(* IEC 61131-3 sources: ZPLC/tools/hil/st_tests, 25 files *)

(* ---- full_language_test.st ---- *)
TYPE State : (INIT, PROCESS, DONE, ERROR); END_TYPE

FUNCTION_BLOCK FB_Logger
    VAR
        LastMsg : WSTRING;
        MsgCount : INT := 0;
    END_VAR

    METHOD PUBLIC Log : BOOL
        VAR_INPUT
            Msg : WSTRING;
        END_VAR
        THIS.LastMsg := Msg;
        THIS.MsgCount := THIS.MsgCount + 1;
        Log := TRUE;
    END_METHOD
END_FUNCTION_BLOCK

FUNCTION_BLOCK FB_Process EXTENDS FB_Logger
    VAR
        Timestamp : DT;
        Result : REAL;
    END_VAR

    METHOD PUBLIC Calc : REAL
        VAR_INPUT
            InVal : REAL;
        END_VAR
        VAR_TEMP
            tmp : REAL;
        END_VAR

        tmp := tmp + InVal * 2.0;
        Calc := tmp;
    END_METHOD
END_FUNCTION_BLOCK

PROGRAM FullTest
    VAR
        machine : FB_Process;
        currentState : State := INIT;

        test_dt : DT;
        calc_res1 AT %QD1 : REAL;
        calc_res2 AT %QD2 : REAL;

        cycle AT %QW0 : INT := 0;

        flag_enum AT %QX12.0 : BOOL;
        flag_oop AT %QX12.1 : BOOL;
        flag_temp AT %QX12.2 : BOOL;
        flag_types AT %QX12.3 : BOOL;
    END_VAR

    cycle := cycle + 1;

    CASE currentState OF
        0: (* INIT *)
            machine.Log(Msg := "Start");
            machine.Timestamp := DT#2024-01-01-12:00:00;
            test_dt := machine.Timestamp;
            currentState := 1;

        1: (* PROCESS *)
            calc_res1 := machine.Calc(InVal := 10.0);
            calc_res2 := machine.Calc(InVal := 20.0);
            currentState := 2;

        2: (* DONE *)
            flag_enum := TRUE;

            IF machine.MsgCount = 1 THEN flag_oop := TRUE; END_IF;

            IF calc_res1 = 20.0 AND calc_res2 = 40.0 THEN flag_temp := TRUE; END_IF;

            IF test_dt > DT#2023-01-01-00:00:00 THEN flag_types := TRUE; END_IF;
    END_CASE;

END_PROGRAM

(* ---- named_params_test.st ---- *)
FUNCTION_BLOCK FB_Calc
    METHOD PUBLIC Add : REAL
        VAR_INPUT
            A : REAL;
            B : REAL;
        END_VAR
        Add := A + B;
    END_METHOD
END_FUNCTION_BLOCK

PROGRAM NamedParamsTest
    VAR
        calc : FB_Calc;
        res AT %QD0 : REAL;
    END_VAR

    res := calc.Add(A := 10.0, B := 20.0);
END_PROGRAM

(* ---- oop_extends.st ---- *)
FUNCTION_BLOCK FB_Base
VAR
    BaseVal : INT;
END_VAR

METHOD PUBLIC InitBase : BOOL
    THIS.BaseVal := 10;
    InitBase := TRUE;
END_METHOD

METHOD PUBLIC GetBase : INT
    GetBase := THIS.BaseVal;
END_METHOD

METHOD PUBLIC VirtualMethod : INT
    VirtualMethod := 111;
END_METHOD
END_FUNCTION_BLOCK

FUNCTION_BLOCK FB_Child EXTENDS FB_Base
VAR
    ChildVal : INT;
END_VAR

METHOD PUBLIC InitChild : BOOL
    THIS.BaseVal := 10;
    THIS.ChildVal := 20;
    InitChild := TRUE;
END_METHOD

METHOD PUBLIC GetChild : INT
    GetChild := THIS.ChildVal;
END_METHOD

METHOD PUBLIC OVERRIDE VirtualMethod : INT
    VirtualMethod := 222;
END_METHOD
END_FUNCTION_BLOCK

PROGRAM TestExtends
VAR
    base : FB_Base;
    child : FB_Child;

    res_base_base : INT;
    res_child_base : INT;
    res_child_child : INT;
    res_virt_base : INT;
    res_virt_child : INT;

    initialized : BOOL := FALSE;
    dummy : BOOL;

    test_passed AT %QX0.0 : BOOL := FALSE;
    debug_val AT %QW1 : INT;
    life_counter AT %QW2 : INT; (* 0x1004 *)
END_VAR

life_counter := life_counter + 1;

IF NOT initialized THEN
    dummy := base.InitBase();
    dummy := child.InitChild();
    initialized := TRUE;
END_IF;

res_base_base := base.GetBase();
res_child_base := child.GetBase();
res_child_child := child.GetChild();

res_virt_base := base.VirtualMethod();
res_virt_child := child.VirtualMethod();

debug_val := res_virt_child;

IF res_base_base = 10 AND
   res_child_base = 10 AND
   res_child_child = 20 AND
   res_virt_base = 111 AND
   res_virt_child = 222 THEN
    test_passed := TRUE;
END_IF;

END_PROGRAM

(* ---- oop_extends_simple.st ---- *)
FUNCTION_BLOCK FB_Base
METHOD PUBLIC GetVal : INT
    GetVal := 111;
END_METHOD
END_FUNCTION_BLOCK

FUNCTION_BLOCK FB_Child EXTENDS FB_Base
METHOD PUBLIC OVERRIDE GetVal : INT
    GetVal := 222;
END_METHOD
END_FUNCTION_BLOCK

PROGRAM SimpleExtends
VAR
    child : FB_Child;
    res : INT;
    debug AT %QW0 : INT;
END_VAR

res := child.GetVal();
debug := res;
END_PROGRAM

(* ---- oop_test.st ---- *)
(*
 * ZPLC OOP HIL Test
 *
 * Tests IEC 61131-3 OOP extensions:
 * - FUNCTION_BLOCK with METHOD
 * - THIS keyword
 * - Method calls on FB instances
 *
 * Memory Layout (OPI starts at 0x1000):
 * - 0x1000: test_passed BOOL
 * - 0x1002: counter_value INT (2 bytes)
 * - 0x1004: method_result INT (2 bytes)
 * - 0x1006: cycle_count INT (2 bytes)
 *)

(* Simple Counter FB with Methods *)
FUNCTION_BLOCK FB_Counter
VAR
    Count : INT;
    MaxVal : INT;
END_VAR

(* Reset counter to zero *)
METHOD PUBLIC Reset : BOOL
    THIS.Count := 0;
    THIS.MaxVal := 100;
    Reset := TRUE;
END_METHOD

(* Increment counter by 1 and return new value *)
METHOD PUBLIC Increment : INT
    THIS.Count := THIS.Count + 1;
    Increment := THIS.Count;
END_METHOD

(* Get current count value *)
METHOD PUBLIC GetValue : INT
    GetValue := THIS.Count;
END_METHOD

(* Add 10 to counter *)
METHOD PUBLIC AddTen : INT
    THIS.Count := THIS.Count + 10;
    AddTen := THIS.Count;
END_METHOD

END_FUNCTION_BLOCK

PROGRAM OOPTest
VAR
    (* Output mappings for test verification *)
    test_passed AT %QX0.0 : BOOL := FALSE;  (* 0x1000 bit 0 *)
    counter_value AT %QW1 : INT;            (* 0x1002 *)
    method_result AT %QW2 : INT;            (* 0x1004 *)
    cycle_count AT %QW3 : INT;              (* 0x1006 *)

    (* FB instance *)
    myCounter : FB_Counter;

    (* Local variables *)
    initialized : BOOL := FALSE;
    temp : INT;
    cycles : INT := 0;
END_VAR

(* Increment cycle counter *)
cycles := cycles + 1;
cycle_count := cycles;

(* Only run initialization once *)
IF NOT initialized THEN
    (* Reset counter to zero *)
    myCounter.Reset();
    initialized := TRUE;
END_IF;

(* Each cycle: increment, then add 10 *)
(* Cycle 1: 0 -> 1 -> 11 *)
(* Cycle 2: 11 -> 12 -> 22 *)

temp := myCounter.Increment();
method_result := myCounter.AddTen();
counter_value := myCounter.GetValue();

(* Test passes if counter >= 11 (at least one full cycle completed) *)
IF counter_value >= 11 THEN
    test_passed := TRUE;
END_IF;

END_PROGRAM

(* ---- user_fb.st ---- *)
FUNCTION_BLOCK MyCounter
VAR_INPUT
    Up : BOOL;
END_VAR
VAR_OUTPUT
    Count : INT := 0;
END_VAR
VAR
    prev_up : BOOL := FALSE;
END_VAR

    (* Rising Edge Detection *)
    IF Up AND NOT prev_up THEN
        Count := Count + 1;
    END_IF;
    prev_up := Up;

END_FUNCTION_BLOCK

PROGRAM UserFBTest
VAR
    c1 : MyCounter;
    clk : BOOL := FALSE;
    res_count AT %QW0 : INT; (* 0x1000 *)

    cycle : INT := 0;
END_VAR

cycle := cycle + 1;

(* Generate pulse every 2 cycles: 0->F, 1->F, 2->T, 3->F, 4->T ... *)
clk := (cycle MOD 2) = 0;

c1(Up := clk);
res_count := c1.Count;

END_PROGRAM

(* ---- vartemp_hil.st ---- *)
FUNCTION_BLOCK FB_TempTest
    METHOD PUBLIC AddTemp : INT
        VAR_INPUT In : INT; END_VAR
        VAR_TEMP tmp : INT := 0; END_VAR

        (* tmp should be 0 at start of every call *)
        tmp := tmp + In;
        AddTemp := tmp;
    END_METHOD
END_FUNCTION_BLOCK

PROGRAM Main
    VAR
        fb : FB_TempTest;
        res1 AT %QW0 : INT;
        res2 AT %QW1 : INT;
    END_VAR

    res1 := fb.AddTemp(In := 10);
    res2 := fb.AddTemp(In := 20);
END_PROGRAM

(* ---- complex_types.st ---- *)
PROGRAM ComplexTypes
VAR
    matrix : ARRAY[0..1, 0..1] OF INT;
    sum : INT;

    (* Result on the output image, byte 0 (0x1000) *)
    res_x AT %QW0 : INT;
END_VAR

(* Initialize Matrix *)
matrix[0,0] := 10;
matrix[0,1] := 20;
matrix[1,0] := 30;
matrix[1,1] := 40;

(* Calculate diagonal sum: 10 + 40 = 50 *)
sum := matrix[0,0] + matrix[1,1];

(* Output *)
res_x := sum;

END_PROGRAM

(* ---- counters_extra.st ---- *)
PROGRAM TestCounters
VAR
    (* CTD Test *)
    myCtd : CTD;
    cd : BOOL;
    ld : BOOL;
    pv : INT := 5;
    q_ctd AT %QX0.0 : BOOL;
    cv_ctd AT %QW1 : INT;

    (* CTUD Test *)
    myCtud : CTUD;
    cu : BOOL;
    cd_ud : BOOL;
    r : BOOL;
    ld_ud : BOOL;
    pv_ud : INT := 5;
    qu AT %QX0.1 : BOOL;
    qd AT %QX0.2 : BOOL;
    cv_ud AT %QW2 : INT;

    step : INT := 0;
    cycles : INT := 0;
END_VAR

cycles := cycles + 1;

(* State Machine to generate edges *)
CASE step OF
    0: (* Init *)
        ld := TRUE; (* CTD: Load 5 *)
        r := TRUE;  (* CTUD: Reset to 0 *)
        step := 1;

    1: (* Release controls *)
        ld := FALSE;
        r := FALSE;
        step := 2;

    2: (* Generate 3 down pulses for CTD *)
        cd := TRUE;
        step := 3;
    3:
        cd := FALSE;
        step := 4;
    4:
        cd := TRUE;
        step := 5;
    5:
        cd := FALSE;
        step := 6;
    6:
        cd := TRUE;
        step := 7;
    7:
        cd := FALSE;
        (* CTD started at 5. 3 pulses -> 2. *)

        (* Generate 6 up pulses for CTUD *)
        cu := TRUE;
        step := 8;
    8:
        cu := FALSE;
        (* Repeat up to 6 times using modulo logic or just linear steps *)
        IF cycles > 30 THEN
            step := 99;
        ELSE
            (* Toggle CU every even/odd step *)
            IF (cycles MOD 2) = 0 THEN cu := TRUE; ELSE cu := FALSE; END_IF;
        END_IF;

    99: (* Done *)
        cu := FALSE;
        cd := FALSE;
END_CASE;

(* Call FBs *)
myCtd(CD := cd, LD := ld, PV := pv);
q_ctd := myCtd.Q;
cv_ctd := myCtd.CV;

myCtud(CU := cu, CD := cd_ud, R := r, LD := ld_ud, PV := pv_ud);
qu := myCtud.QU;
qd := myCtud.QD;
cv_ud := myCtud.CV;

END_PROGRAM

(* ---- loop_control.st ---- *)
PROGRAM LoopControl
VAR
    i : INT;
    j : INT;
    sum : INT := 0;

    res_exit AT %QW0 : INT;    (* 0x1000 *)
    res_cont AT %QW1 : INT;    (* 0x1002 *)
END_VAR

(* EXIT Test: Stop at 5 *)
FOR i := 1 TO 10 DO
    IF i = 5 THEN
        EXIT;
    END_IF;
END_FOR;
res_exit := i;

(* CONTINUE Test: Sum all except 3 (1+2+4+5=12) *)
sum := 0;
FOR j := 1 TO 5 DO
    IF j = 3 THEN
        CONTINUE;
    END_IF;
    sum := sum + j;
END_FOR;
res_cont := sum;

END_PROGRAM

(* ---- loop_test.st ---- *)
PROGRAM LoopTest
VAR
    i : INT := 0;
    j : INT := 0;

    res_while AT %QW0 : INT;  (* 0x1000 *)
    res_repeat AT %QW1 : INT; (* 0x1002 *)
END_VAR

(* WHILE Loop *)
WHILE i < 10 DO
    i := i + 1;
END_WHILE;
res_while := i;

(* REPEAT Loop *)
REPEAT
    j := j + 1;
UNTIL j = 20
END_REPEAT;
res_repeat := j;

(* Reset for next cycle *)
IF i >= 10 THEN i := 0; END_IF;
IF j >= 20 THEN j := 0; END_IF;

END_PROGRAM

(* ---- master_blinky.st ---- *)
PROGRAM MasterBlinky
VAR
    fast_tmr : TON;
    slow_tmr : TON;

    fast_state AT %QX0.1 : BOOL; (* GP1 *)
    slow_state AT %QX0.0 : BOOL; (* GP0 *)

    cycle_count : INT := 0;
END_VAR

(* Fast Blinky (100ms ON / 100ms OFF) *)
fast_tmr(IN := NOT fast_tmr.Q, PT := T#100ms);
IF fast_tmr.Q THEN
    fast_state := NOT fast_state;
END_IF;

(* Slow Blinky (500ms ON / 500ms OFF) *)
slow_tmr(IN := NOT slow_tmr.Q, PT := T#500ms);
IF slow_tmr.Q THEN
    slow_state := NOT slow_state;
END_IF;

cycle_count := cycle_count + 1;

END_PROGRAM

(* ---- master_math_control.st ---- *)
PROGRAM MathControlTest
VAR
    (* Math Results *)
    res_sqrt AT %QD1 : REAL;   (* 0x1004 *)
    res_ln AT %QD2 : REAL;     (* 0x1008 *)
    res_sin AT %QD3 : REAL;   (* 0x100C *)
    res_expt AT %QW8 : INT;   (* 0x1010 *)

    (* Control Results *)
    res_for AT %QW9 : INT;    (* 0x1012 *)
    res_case AT %QW10 : INT;   (* 0x1014 *)

    (* Internal vars *)
    i : INT;
    temp_sum : INT := 0;
    case_sel : INT := 2;
END_VAR

(* 1. Math Tests *)
res_sqrt := SQRT(2.0);
res_ln := LN(2.7182818);
res_sin := SIN(1.570796);
res_expt := REAL_TO_INT(EXPT(2.0, 8));

(* 2. FOR loop test *)
temp_sum := 0;
FOR i := 1 TO 10 DO
    temp_sum := temp_sum + i;
END_FOR;
res_for := temp_sum;

(* 3. CASE test *)
CASE case_sel OF
    1: res_case := 10;
    2: res_case := 20;
    3: res_case := 30;
ELSE
    res_case := 99;
END_CASE;

END_PROGRAM

(* ---- master_test.st ---- *)
PROGRAM MasterTest
VAR
    test_cycle : INT := 0;
    latch_rs : RS;
    latch_sr : SR;
    trig_r : R_TRIG;
    counter : CTU;

    res_rs AT %QX0.0 : BOOL;
    res_sr AT %QX0.1 : BOOL;
    res_trig AT %QX0.2 : BOOL;
    res_ctu AT %QX0.3 : BOOL;
END_VAR

test_cycle := test_cycle + 1;

(* 1. Test RS: Set once and keep it *)
latch_rs(S := (test_cycle = 5), R1 := FALSE);
res_rs := latch_rs.Q1;

(* 2. Test SR: Set once and keep it *)
latch_sr(S1 := (test_cycle = 5), R := FALSE);
res_sr := latch_sr.Q1;

(* 3. Test Trigger: Pulse and latch the result *)
trig_r(CLK := (test_cycle = 5));
IF trig_r.Q THEN
    res_trig := TRUE;
END_IF;

(* 4. Test Counter: Count to 5 and stay there *)
counter(CU := (test_cycle <= 10 AND (test_cycle MOD 2 = 0)), PV := 5, R := (test_cycle = 1));
res_ctu := counter.Q;

END_PROGRAM

(* ---- master_test_2.st ---- *)
PROGRAM MasterTest2
VAR
    test_cycle : INT := 0;
    timer_off : TOF;
    timer_pulse : TP;
    i : INT;
    sum : INT := 0;
    case_val : INT := 0;

    (* Results on the output image: STOP puts the outputs in their safe state, so they are read while it runs *)
    res_tof AT %QX0.0 : BOOL;
    res_tp AT %QX0.1 : BOOL;
    res_for AT %QW1 : INT;
    res_case AT %QW2 : INT;
END_VAR

test_cycle := test_cycle + 1;

timer_off(IN := (test_cycle = 5), PT := T#500ms);
IF test_cycle = 10 AND timer_off.Q THEN
    res_tof := TRUE;
END_IF;

timer_pulse(IN := (test_cycle = 5), PT := T#500ms);
IF test_cycle = 7 AND timer_pulse.Q THEN
    res_tp := TRUE;
END_IF;

IF test_cycle = 10 THEN
    sum := 0;
    FOR i := 1 TO 5 DO
        sum := sum + i;
    END_FOR;
    res_for := sum;
END_IF;

IF test_cycle = 10 THEN
    case_val := 2;
    CASE case_val OF
        1: res_case := 100;
        2: res_case := 200;
    ELSE
        res_case := 0;
    END_CASE;
END_IF;

END_PROGRAM

(* ---- math_real.st ---- *)
PROGRAM MathReal
VAR
    angles : ARRAY[0..2] OF REAL;
    sines : ARRAY[0..2] OF REAL;
    i : INT;

    (* OPI Layout: *)
    (* 0x1000: result_ok (INT, 2 bytes) *)
    (* 0x1004: debug_val (REAL, 4 bytes) *)

    result_ok AT %QW0 : INT;
    debug_val AT %QD1 : REAL;
END_VAR

angles[0] := 0.0;
angles[1] := 1.570796;
angles[2] := 3.141592;

FOR i := 0 TO 2 DO
    sines[i] := SIN(angles[i]);
END_FOR;

(* Store result for debugging *)
debug_val := sines[1];

IF sines[1] > 0.99 AND sines[1] < 1.01 THEN
    result_ok := 1;
ELSE
    result_ok := 0;
END_IF;

END_PROGRAM

(* ---- moving_avg.st ---- *)
PROGRAM MovingAvg
VAR
    buffer : ARRAY[0..4] OF INT;
    i : INT;
    sum : DINT;
    avg AT %QW0 : INT; (* Result at 0x1000 *)

    raw_val : INT := 0;
    counter : INT := 0;
END_VAR

(* Simulate Input *)
counter := counter + 10;
IF counter > 100 THEN
    counter := 0;
END_IF;
raw_val := counter;

(* Shift Buffer (Unrolled to avoid negative step compiler bug) *)
buffer[4] := buffer[3];
buffer[3] := buffer[2];
buffer[2] := buffer[1];
buffer[1] := buffer[0];

(* Insert new value *)
buffer[0] := raw_val;

(* Calculate Average *)
sum := 0;
FOR i := 0 TO 4 DO
    (* Implicit conversion INT to DINT is handled by VM stack *)
    sum := sum + buffer[i];
END_FOR;

(* Implicit conversion DINT to INT *)
avg := sum / 5;

END_PROGRAM

(* ---- pointer_test.st ---- *)
PROGRAM PointerTest
VAR
    val : INT;
    ptr : REF_TO INT;

    res_read AT %QW0 : INT; (* 0x1000 *)
    res_write AT %QW1 : INT; (* 0x1002 *)
END_VAR

(* Initialize val each cycle to verify read before write *)
val := 42;

(* 1. Reference *)
ptr := REF(val);

(* 2. Dereference Read *)
res_read := ptr^;

(* 3. Dereference Write *)
ptr^ := 99;
res_write := val;

END_PROGRAM

(* ---- process_test.st ---- *)
PROGRAM ProcessTest
VAR
    (* --- HYSTERESIS Test --- *)
    hyst : HYSTERESIS;
    hyst_in : REAL;
    hyst_q AT %QX0.0 : BOOL;

    (* --- DEADBAND Test --- *)
    db : DEADBAND;
    db_in : REAL := 10.0;
    db_out : REAL;

    (* --- LAG_FILTER Test --- *)
    lag : LAG_FILTER;
    lag_in : REAL := 100.0;
    lag_out AT %QD1 : REAL;

    (* --- RAMP_REAL Test --- *)
    ramp : RAMP_REAL;
    ramp_in : REAL := 50.0;
    ramp_out : REAL;

    (* --- PID Test --- *)
    pid : PID_Compact;
    pid_sp : REAL := 10.0;
    pid_pv : REAL := 0.0;
    pid_out AT %QD2 : REAL;

    cycle : INT := 0;
END_VAR

cycle := cycle + 1;

(* 1. HYSTERESIS: High=10, Low=5. Input sweeps *)
IF cycle < 5 THEN
    hyst_in := 0.0;
ELSIF cycle < 10 THEN
    hyst_in := 12.0; (* > High, Q -> TRUE *)
ELSIF cycle < 15 THEN
    hyst_in := 8.0;  (* < High but > Low, Q stays TRUE *)
ELSE
    hyst_in := 2.0;  (* < Low, Q -> FALSE *)
END_IF;

hyst(IN := hyst_in, HIGH := 10.0, LOW := 5.0);
hyst_q := hyst.Q;

(* 2. DEADBAND: Width=2.0. Input changes *)
(* Default db_out starts at 0? No, internal state init 0 *)
IF cycle > 5 THEN db_in := 11.5; END_IF; (* diff 1.5 < 2, should ignore? Wait, ref is _last *)
IF cycle > 10 THEN db_in := 13.0; END_IF; (* diff vs last update *)

db(IN := db_in, WIDTH := 2.0);
db_out := db.OUT;

(* 3. LAG_FILTER: Input step 0->100. Gain 0.1 *)
(* Output should approach 100 exponentially *)
lag(IN := lag_in, GAIN := 0.1);
lag_out := lag.OUT;

(* 4. RAMP_REAL: Input step 0->50. Rate 1.0 per cycle *)
(* Output should increase by 1.0 each cycle *)
ramp(IN := ramp_in, RATE := 1.0);
ramp_out := ramp.OUT;

(* 5. PID: SP=10, PV=0. P-only first (KI=0, KD=0) *)
(* Error=10. KP=2.0 -> Out=20.0 *)
pid(SP := pid_sp, PV := pid_pv, KP := 2.0, KI := 0.0, KD := 0.0, DT := 0.1, OUT_MIN := -100.0, OUT_MAX := 100.0);
pid_out := pid.OUT;

END_PROGRAM

(* ---- struct_revisited.st ---- *)
TYPE
    Point : STRUCT
        x : INT;
        y : INT;
    END_STRUCT;
END_TYPE

PROGRAM StructTest
VAR
    p1 : Point;
    sum AT %QW0 : INT; (* 0x1000 *)
END_VAR

p1.x := 10;
p1.y := 20;
sum := p1.x + p1.y;

END_PROGRAM

(* ---- struct_test.st ---- *)
TYPE
    MyPoint : STRUCT
        x : INT;
        y : INT;
    END_STRUCT;
END_TYPE

PROGRAM StructTest
VAR
    p1 : MyPoint;
    sum AT %QW0 : INT; (* 0x1000 *)
END_VAR

p1.x := 10;
p1.y := 20;
sum := p1.x + p1.y;

END_PROGRAM

(* ---- test_ctu.st ---- *)
PROGRAM TestCTU
VAR
    count1 : CTU;
    clk : BOOL := TRUE;
    out_full AT %QX0.0 : BOOL;
    cv AT %QW1 : INT;
END_VAR

count1(CU := clk, PV := 5, R := FALSE);
out_full := count1.Q;
cv := count1.CV;

clk := NOT clk;
END_PROGRAM

(* ---- test_rs.st ---- *)
PROGRAM TestRS
VAR
    latch : RS;
    s_in AT %IX0.0 : BOOL;
    r_in AT %IX0.1 : BOOL;
    q_out AT %QX0.0 : BOOL;
END_VAR

latch(S := s_in, R1 := r_in);
q_out := latch.Q1;

END_PROGRAM

(* ---- test_ton.st ---- *)
PROGRAM TestTON
VAR
    timer1 : TON;
    out1 AT %QX0.0 : BOOL;
    et AT %QD1 : TIME;
END_VAR

timer1(IN := TRUE, PT := T#200ms);
out1 := timer1.Q;
et := timer1.ET;
END_PROGRAM

(* ---- user_function.st ---- *)
FUNCTION Hypotenuse : REAL
VAR_INPUT
    a : REAL;
    b : REAL;
END_VAR
    Hypotenuse := SQRT(a*a + b*b);
END_FUNCTION

PROGRAM UserFuncTest
VAR
    res AT %QD0 : REAL; (* 0x1000 *)
    cycle AT %QW2 : INT; (* 0x1004 *)
    counter : INT := 0;
END_VAR

counter := counter + 1;
cycle := counter;

res := Hypotenuse(3.0, 4.0);

END_PROGRAM
